// TIA Portal V20 export
// export: Created 2026-11-20T10:15:00.000Z, ExportSetting WithDefaults
FUNCTION_BLOCK "FB_Conveyor"   // FB12, LAD
TITLE = Belt conveyor
{ S7_Optimized_Access := 'TRUE' }
AUTHOR : controls
VERSION : 0.2
// stored: AutoNumber true, SetENOAutomatically false
   VAR_INPUT
      Start : Bool;   // Start push button
      Stop : Bool;   // Stop push button (NC)
      Jam : Bool;   // Jam photo-eye blocked
   END_VAR
   VAR_OUTPUT
      Run : Bool;
      JamAlarm : Bool;
   END_VAR
   VAR
      JamTimer : IEC_TIMER;
      Speed : Real := 1.5;
   END_VAR
BEGIN

REGION Network 1: Run latch
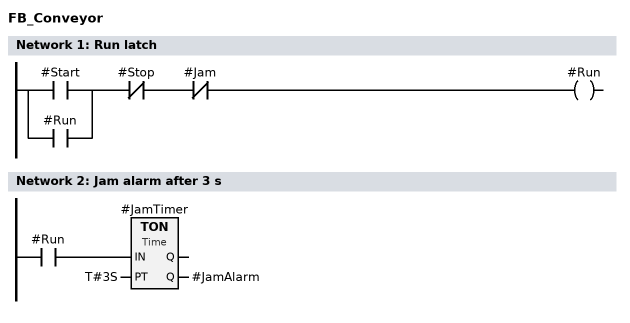
   #Run := (#Start OR #Run) AND NOT #Stop AND NOT #Jam;
END_REGION

REGION Network 2: Jam alarm after 3 s
   RUNG wire#powerrail
      Contact( #Run )
      { S7_Templates := "time_type := Time" } #JamTimer.TON(pt := T#3S, q => #JamAlarm)
   END_RUNG
   // the same network as SCL:
   #JamTimer.TON(IN := #Run, PT := T#3S, Q => #JamAlarm);
END_REGION
END_FUNCTION_BLOCK
